Fanuc KAREL source: kx00012.KL

-- PROVISIONAL review KL for V1013-1; original PC SHA256 87d39c06785eeb930a5310ec7d97cb7ffa47c09408d1999c624883f28ae54e0e
-- Incomplete behavior may be omitted. Consult companion uncertainty JSON. Do not deploy.
PROGRAM KX00012
%NOLOCKGROUP
VAR
  I : INTEGER
  J : INTEGER
  B : BOOLEAN
  F : FILE
  S : STRING[80]
-- UNRESOLVED_DECL P type=000102
BEGIN
  -- UNRESOLVED_PC offsets 5-7; opcodes 9C,66
  -- UNRESOLVED_PC offsets 12-16; opcodes 7F
END KX00012
